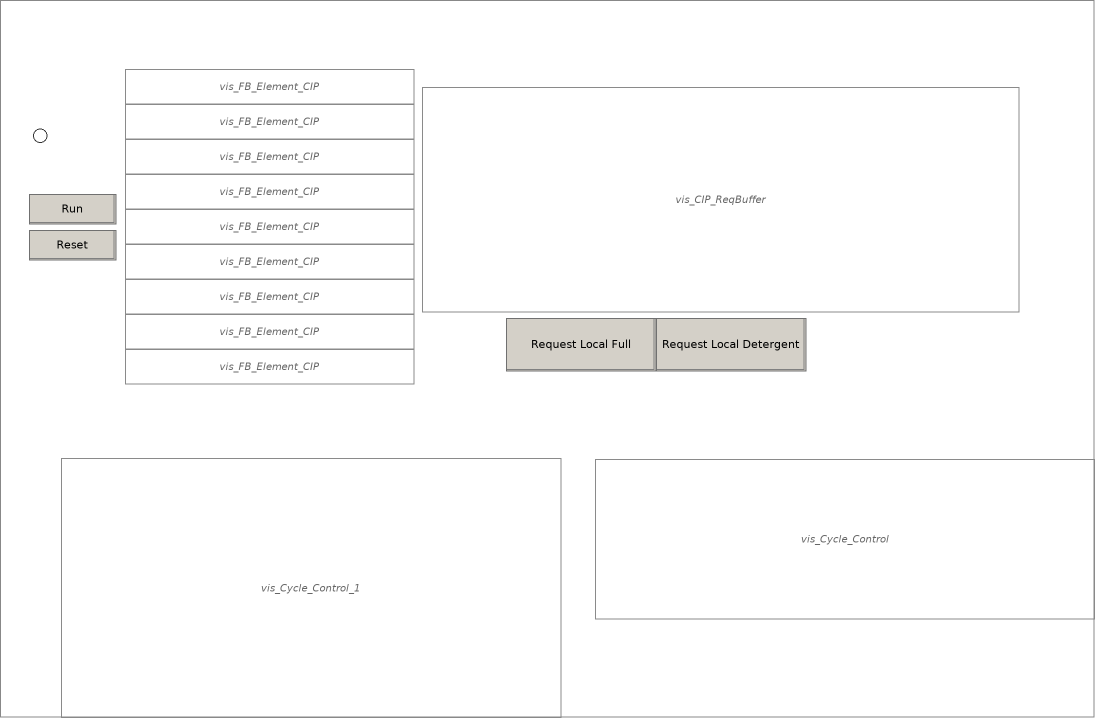
VISUALIZATION vis_CIP  // 1095x718
    Button (29,194 87x30), "Run", colour toggle: fbCIP.bRun
        toggle fbCIP.bRun
    Button (29,230 87x30), "Reset", colour toggle: fbCIP.SFCReset
        toggle fbCIP.SFCReset
    Button (506,318 150x53), "Request Local Full"
        tap fbCIP.rtReqLocalCIP_Full_HMI.CLK
    Button (656,318 150x53), "Request Local Detergent"
        tap fbCIP.rtReqLocalCIP_Detergent_HMI.CLK
    RadioButton (31,86 102x99), variable: fbCIP.eMode
        Areas[0]: Text=Off
        Areas[1]: Text=Manual
        Areas[2]: Text=Auto
    Frame (422,87 597x225)
        shows vis_CIP_ReqBuffer()
    Group (125,69 289x315)
        Frame (0,0 289x35)
            shows vis_FB_Element_CIP(fb := fbElement[E_Element_List.eTank_1])
        Frame (0,35 289x35)
            shows vis_FB_Element_CIP(fb := fbElement[E_Element_List.eTank_2])
        Frame (0,70 289x35)
            shows vis_FB_Element_CIP(fb := fbElement[E_Element_List.eTank_3])
        Frame (0,105 289x35)
            shows vis_FB_Element_CIP(fb := fbElement[E_Element_List.eTank_4])
        Frame (0,140 289x35)
            shows vis_FB_Element_CIP(fb := fbElement[E_Element_List.eTriBlender_Marinada])
        Frame (0,175 289x35)
            shows vis_FB_Element_CIP(fb := fbElement[E_Element_List.eTriBlender_Color])
        Frame (0,210 289x35)
            shows vis_FB_Element_CIP(fb := fbElement[E_Element_List.eLine_Marinada])
        Frame (0,245 289x35)
            shows vis_FB_Element_CIP(fb := fbElement[E_Element_List.eLine_Color])
        Frame (0,280 289x35)
            shows vis_FB_Element_CIP(fb := fbCIP.fbElement_Blank)
    Frame (595,459 500x160)
        shows vis_Cycle_Control(fb := fbCIP, sName := 'CIP')
    Frame (61,458 500x260)
        shows vis_Cycle_Control_1(fb := fbCIP, sName := 'CIP')
END_VISUALIZATION

(* stored: Version 1.1.0.1, ProductVersion 3.1.4024.12
   Visu vis_CIP: Id {0d0580f4-81f0-46fe-86ed-d2fa56eb530d} *)
